Fanuc KAREL source: kx00028.KL

-- PROVISIONAL review KL for V1013-1; original PC SHA256 c9e804f80e005fe72b9530c371b9ab84f3a23fbc319ae98cc3622e0ed91d7398
-- Incomplete behavior may be omitted. Consult companion uncertainty JSON. Do not deploy.
PROGRAM KX00028
%NOLOCKGROUP
VAR
  I : INTEGER
  J : INTEGER
  B : BOOLEAN
  F : FILE
  S : STRING[80]
-- UNRESOLVED_DECL P type=000102
BEGIN
  -- UNRESOLVED_PC offsets 5-12; opcodes 9D,23
  -- UNRESOLVED_PC offsets 17-21; opcodes 7F
END KX00028
